Fanuc KAREL source: kb00050.KL

-- PROVISIONAL review KL for V770-1; original PC SHA256 a69ff8e11f059c000d38095b178f56f6f3843b116b1de77bdcf2819e49a0e7c9
-- Incomplete behavior may be omitted. Consult companion uncertainty JSON. Do not deploy.
PROGRAM KB00050
%NOLOCKGROUP
BEGIN
  -- UNRESOLVED_PC offsets 5-14; opcodes 3F,75
  -- UNRESOLVED_PC offsets 19-28; opcodes 3F,75
  -- UNRESOLVED_PC offsets 33-42; opcodes 3F,75
  -- UNRESOLVED_PC offsets 47-56; opcodes 3F,75
  -- UNRESOLVED_PC offsets 61-68; opcodes 9D,23
  -- UNRESOLVED_PC offsets 73-80; opcodes 9D,23
  -- UNRESOLVED_PC offsets 85-92; opcodes 9D,23
  -- UNRESOLVED_PC offsets 97-104; opcodes 9D,23
  -- UNRESOLVED_PC offsets 109-116; opcodes 9D,23
  -- UNRESOLVED_PC offsets 121-189; opcodes 27,22,2A,22,2A,22,2A,22,2A,22,22,22,22,22,27,9D,31
  -- UNRESOLVED_PC offsets 194-198; opcodes 7F
END KB00050
